(* PLC project FillingLine, Jack Lai Filling line training bench 0.1 *)
(* stored: creationDateTime 2026-11-03T12:00:00 *)

PROGRAM FillingLine
  VAR_INPUT
    Start AT %IX0.0 : BOOL;
    Stop AT %IX0.1 : BOOL;
    Reset AT %IX0.2 : BOOL;
    EStopOK AT %IX0.3 : BOOL;
    GuardClosed AT %IX0.4 : BOOL;
    TankOK AT %IX0.5 : BOOL;
    BottleAtFill AT %IX0.6 : BOOL;
    ExitSensor AT %IX0.7 : BOOL;
    JamSwitch AT %IX1.0 : BOOL;
  END_VAR
  VAR_OUTPUT
    Run AT %QX0.0 : BOOL;
    Conveyor AT %QX0.1 : BOOL;
    Valve AT %QX0.2 : BOOL;
    Alarm AT %QX0.3 : BOOL;
    BatchDone AT %QX0.4 : BOOL;
    FillBlocked AT %QX0.5 : BOOL;
  END_VAR
  VAR
    Fault : BOOL;
    Filled : BOOL;
    StartEdge : R_TRIG;
    ExitEdge : R_TRIG;
    BatchCount : CTU;
    JamTimer : TON;
    FillTimer : TON;
    FillClearTimer : TON;
  END_VAR

(* LD diagram, written out as Structured Text *)
StartEdge(CLK := Start);
ExitEdge(CLK := ExitSensor);
BatchCount(CU := ExitEdge.Q AND Run, R := Reset, PV := 5);
JamTimer(IN := Conveyor AND NOT ExitSensor, PT := T#3000ms);
FillClearTimer(IN := Run AND Filled AND BottleAtFill, PT := T#1000ms);
FillTimer(IN := Run AND BottleAtFill AND NOT Filled, PT := T#1000ms);
FillBlocked := FillClearTimer.Q OR FillBlocked AND NOT Reset OR FillBlocked AND BottleAtFill;
Fault := NOT EStopOK OR NOT GuardClosed OR NOT TankOK OR JamSwitch OR JamTimer.Q OR Stop AND Run AND BottleAtFill AND NOT Filled OR Fault AND NOT Reset OR Fault AND BottleAtFill OR FillBlocked;
Run := (StartEdge.Q OR Run) AND NOT Stop AND EStopOK AND GuardClosed AND TankOK AND NOT Fault AND NOT BatchCount.Q;
Filled := (FillTimer.Q OR Filled) AND BottleAtFill AND Run;
Conveyor := Run AND (NOT BottleAtFill OR Filled);
Valve := Run AND BottleAtFill AND NOT Filled;
Alarm := Fault;
BatchDone := BatchCount.Q;
END_PROGRAM

CONFIGURATION LineConfig
  RESOURCE CPU ON PLC
    TASK Scan(INTERVAL := T#50ms, PRIORITY := 0);
    PROGRAM Line WITH Scan : FillingLine;
  END_RESOURCE
END_CONFIGURATION
